(* Logix 5000 project; controller CIP_14485201 vendor 1 type 14 code 216 rev 38.11; software revision 38.01; part 4 of 12 *)
(* tags used below, declared in another part *)
   Alarm_Ack : INT[8];   // ALARMS ACKNOWLEDGE BITS
   Alarm_Present : INT[8];   // ALARM MSGS 1-127 PRESENT BITS
   Alarm_Remote_Ack_All : BOOL;   // SYSTEM ALARM ACK ALL TAG USED ON ALARM SETUP ADVANCED TAB TOGGLES EVEYTIME THE ACK_ALL BUTTON IS PUSHED
   Alarm_Timer : TIMER[128];   // ALARM MSGS 1-127 DELAY TIMERS
   Bit : BOOL[128];   // BIT
   IO_Status : INT;   // REMOTE I/O STATUS
   IO_Status_Masked : INT;   // REMOTE I/O STATUS MASK
   OpCode_Pin : DINT[5];   // OPCODE PIN ARRAY
   Process_Heartbeat_Memory : BOOL;
   Process_to_CIP : Process_to_CIP;   // PROCESS SIGNALS TO CIP
   Recipe : RECIPE[41];   // RECIPES
   SCLD_DrainValve_Feedback : SCALE;   // DRAIN FLOW FEEDBACK POSITION 0-100%
   SCLD_Supply_Flow : SCALE;   // SUPPLY FLOW 0-60 GPM
   SCLD_Supply_Press : SCALE;   // SUPPLY PRESSURE 0-100 PSIG
   SCLD_Supply_Temp : SCALE;   // SUPPLY TEMPERATURE 0-100°C
   SCLD_SupplyValve_Feedback : SCALE;   // SUPPLY FLOW FEEDBACK POSITION 0-100%
   SP_DrainValve_HighDeadband : REAL;   // CURRENT DRAIN VALVE DEADBAND SETPOINT
   SP_DrainValve_LowDeadband : REAL;   // CURRENT DRAIN VALVE DEADBAND SETPOINT
   SP_SupplyValve_HighDeadband : REAL;   // CURRENT SUPPLY VALVE DEADBAND SETPOINT
   SP_SupplyValve_LowDeadband : REAL;   // CURRENT SUPPLY VALVE DEADBAND SETPOINT
   Timer : TIMER[99];   // TIMER
   Timer_Chem1_Pump : TIMER[7];   // CHEM #1 CONTROL TIMERS
   Timer_Chem2_Pump : TIMER[7];   // CHEM #2 CONTROL TIMERS
(* MainProgram, continued *)

ROUTINE _05_ALARMS   (* ladder *)
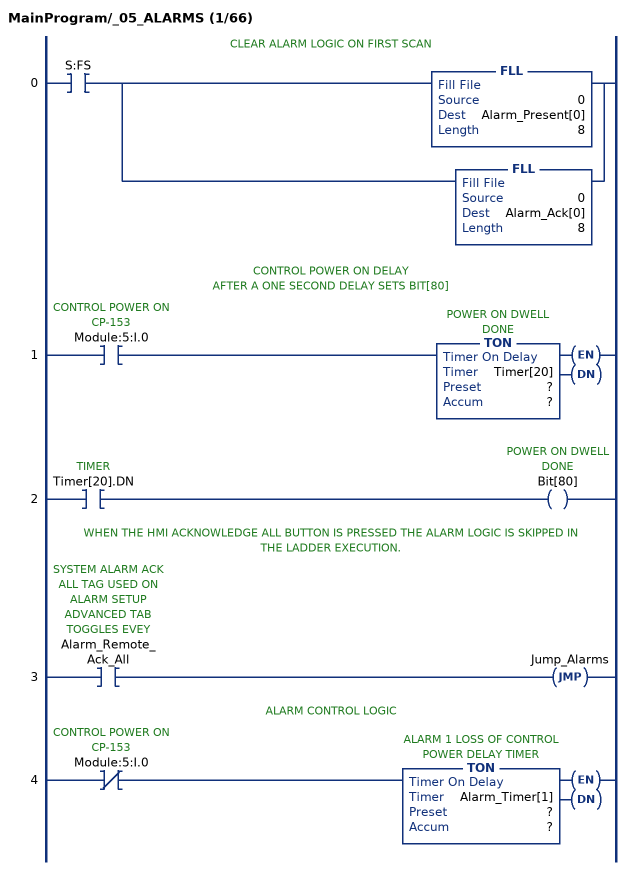
   // CLEAR ALARM LOGIC ON FIRST SCAN
   0: XIC(S:FS)[FLL(0,Alarm_Present[0],8) ,FLL(0,Alarm_Ack[0],8) ];
   // CONTROL POWER ON DELAY
   // AFTER A ONE SECOND DELAY SETS BIT[80]
   1: XIC(Module:5:I.0)TON(Timer[20],?,?);
   2: XIC(Timer[20].DN)OTE(Bit[80]);
   // WHEN THE HMI ACKNOWLEDGE ALL BUTTON IS PRESSED THE ALARM LOGIC IS SKIPPED IN THE LADDER EXECUTION.
   3: XIC(Alarm_Remote_Ack_All)JMP(Jump_Alarms);
   // ALARM CONTROL LOGIC
   4: XIO(Module:5:I.0)TON(Alarm_Timer[1],?,?);
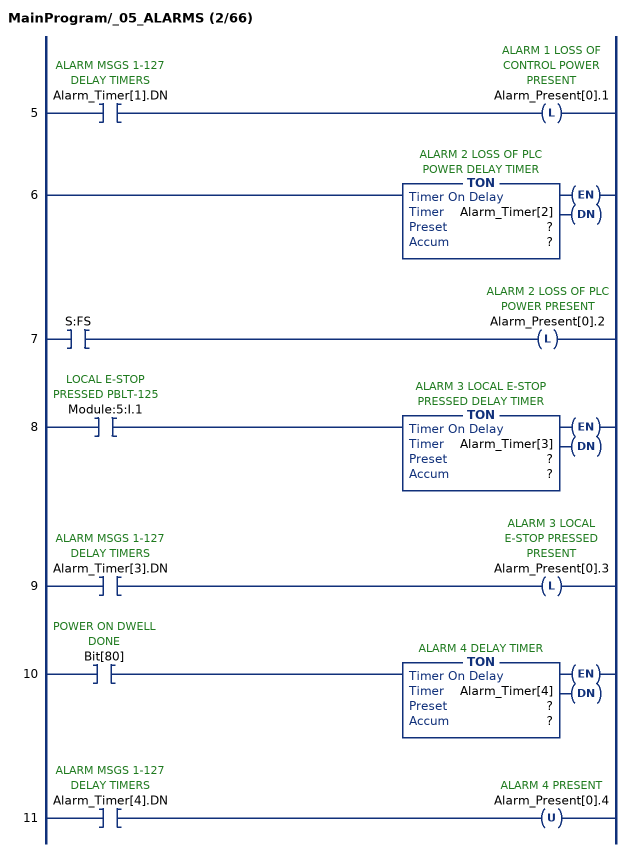
   5: XIC(Alarm_Timer[1].DN)OTL(Alarm_Present[0].1);
   6: TON(Alarm_Timer[2],?,?);
   7: XIC(S:FS)OTL(Alarm_Present[0].2);
   8: XIC(Module:5:I.1)TON(Alarm_Timer[3],?,?);
   9: XIC(Alarm_Timer[3].DN)OTL(Alarm_Present[0].3);
   10: XIC(Bit[80])TON(Alarm_Timer[4],?,?);
   11: XIC(Alarm_Timer[4].DN)OTU(Alarm_Present[0].4);
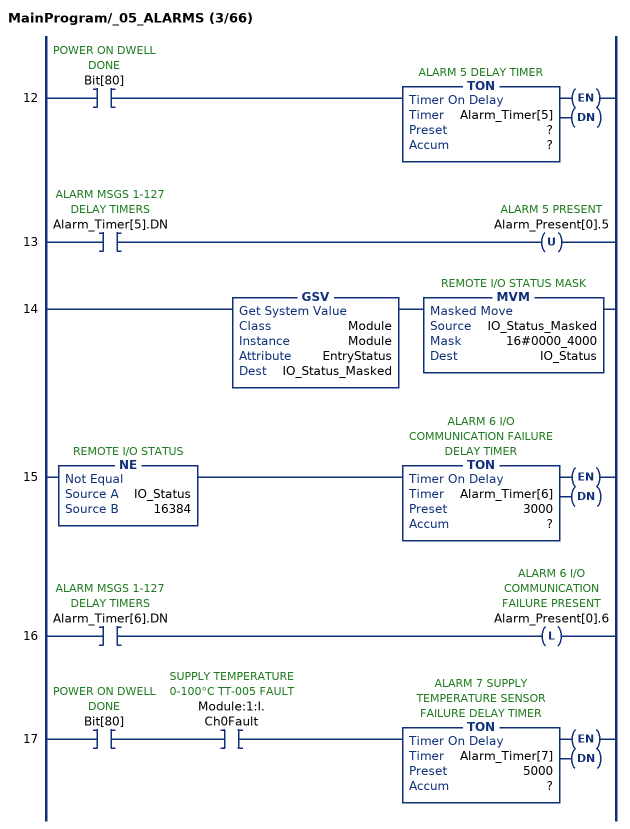
   12: XIC(Bit[80])TON(Alarm_Timer[5],?,?);
   13: XIC(Alarm_Timer[5].DN)OTU(Alarm_Present[0].5);
   14: GSV(Module,Module,EntryStatus,IO_Status_Masked)MVM(IO_Status_Masked,16#0000_4000,IO_Status);
   15: NE(IO_Status,16384)TON(Alarm_Timer[6],?,?);
   16: XIC(Alarm_Timer[6].DN)OTL(Alarm_Present[0].6);
   17: XIC(Bit[80])XIC(Module:1:I.Ch0Fault)TON(Alarm_Timer[7],?,?);
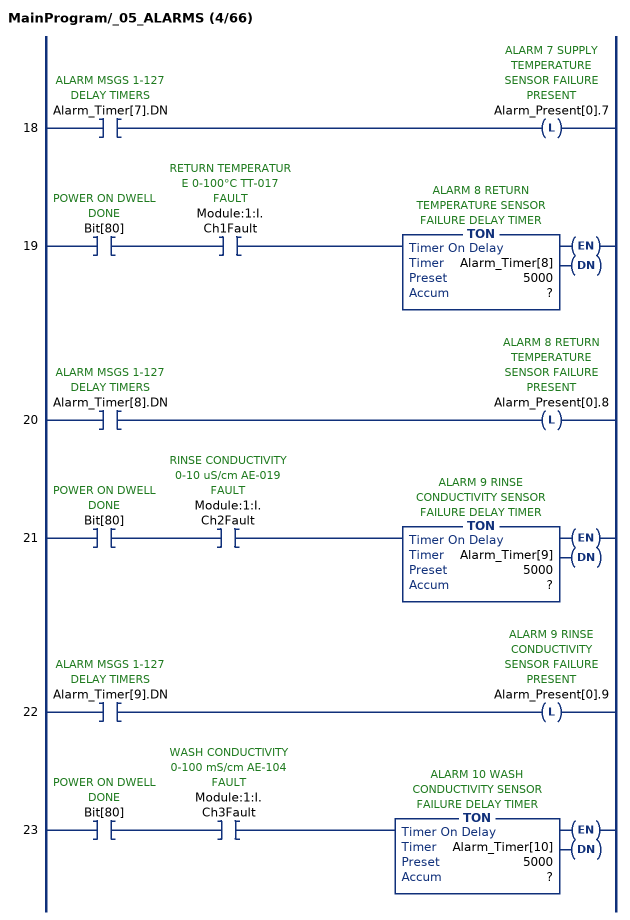
   18: XIC(Alarm_Timer[7].DN)OTL(Alarm_Present[0].7);
   19: XIC(Bit[80])XIC(Module:1:I.Ch1Fault)TON(Alarm_Timer[8],?,?);
   20: XIC(Alarm_Timer[8].DN)OTL(Alarm_Present[0].8);
   21: XIC(Bit[80])XIC(Module:1:I.Ch2Fault)TON(Alarm_Timer[9],?,?);
   22: XIC(Alarm_Timer[9].DN)OTL(Alarm_Present[0].9);
   23: XIC(Bit[80])XIC(Module:1:I.Ch3Fault)TON(Alarm_Timer[10],?,?);
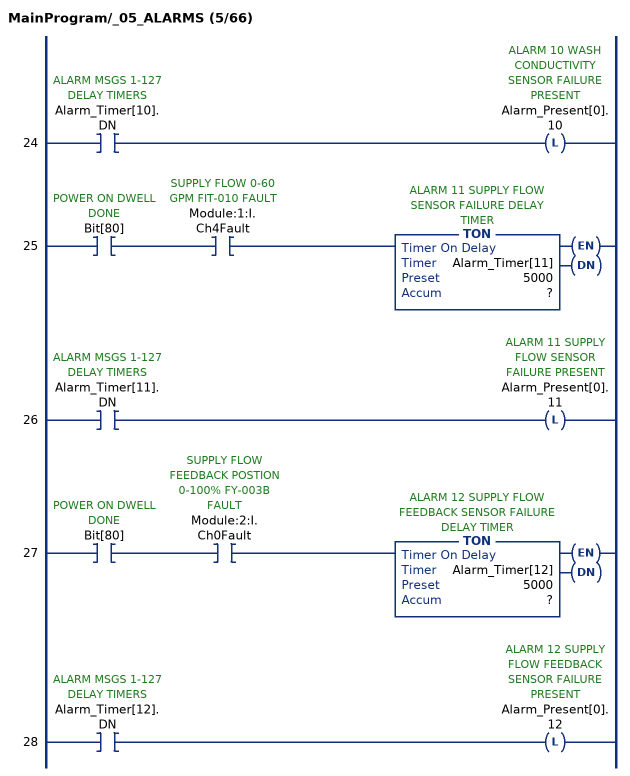
   24: XIC(Alarm_Timer[10].DN)OTL(Alarm_Present[0].10);
   25: XIC(Bit[80])XIC(Module:1:I.Ch4Fault)TON(Alarm_Timer[11],?,?);
   26: XIC(Alarm_Timer[11].DN)OTL(Alarm_Present[0].11);
   27: XIC(Bit[80])XIC(Module:2:I.Ch0Fault)TON(Alarm_Timer[12],?,?);
   28: XIC(Alarm_Timer[12].DN)OTL(Alarm_Present[0].12);
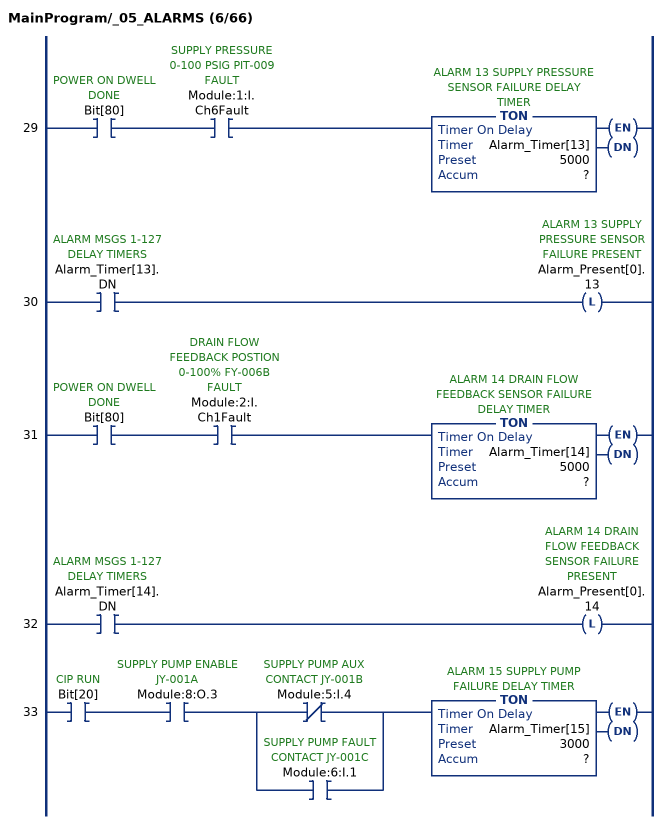
   29: XIC(Bit[80])XIC(Module:1:I.Ch6Fault)TON(Alarm_Timer[13],?,?);
   30: XIC(Alarm_Timer[13].DN)OTL(Alarm_Present[0].13);
   31: XIC(Bit[80])XIC(Module:2:I.Ch1Fault)TON(Alarm_Timer[14],?,?);
   32: XIC(Alarm_Timer[14].DN)OTL(Alarm_Present[0].14);
   33: XIC(Bit[20])XIC(Module:8:O.3)[XIO(Module:5:I.4) ,XIC(Module:6:I.1) ]TON(Alarm_Timer[15],?,?);
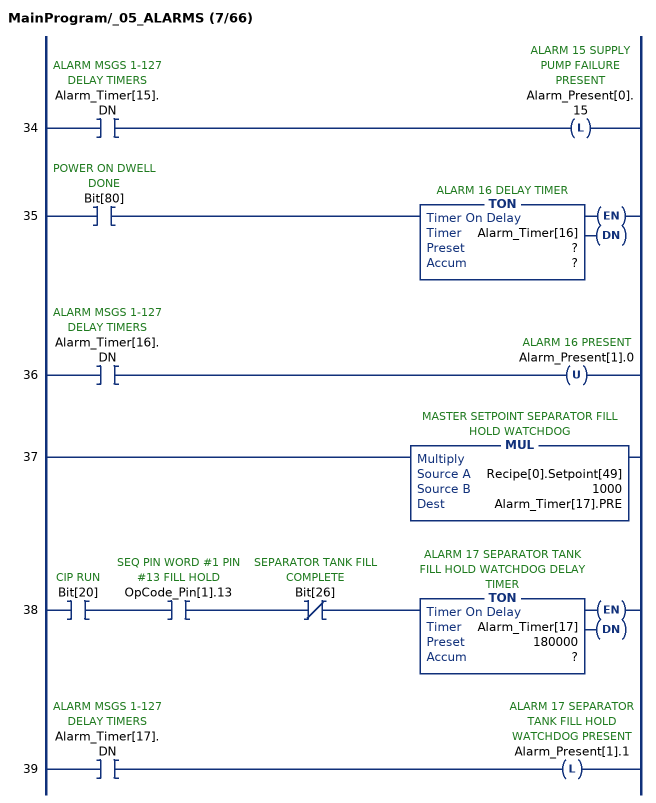
   34: XIC(Alarm_Timer[15].DN)OTL(Alarm_Present[0].15);
   35: XIC(Bit[80])TON(Alarm_Timer[16],?,?);
   36: XIC(Alarm_Timer[16].DN)OTU(Alarm_Present[1].0);
   37: MUL(Recipe[0].Setpoint[49],1000,Alarm_Timer[17].PRE);
   38: XIC(Bit[20])XIC(OpCode_Pin[1].13)XIO(Bit[26])TON(Alarm_Timer[17],?,?);
   39: XIC(Alarm_Timer[17].DN)OTL(Alarm_Present[1].1);
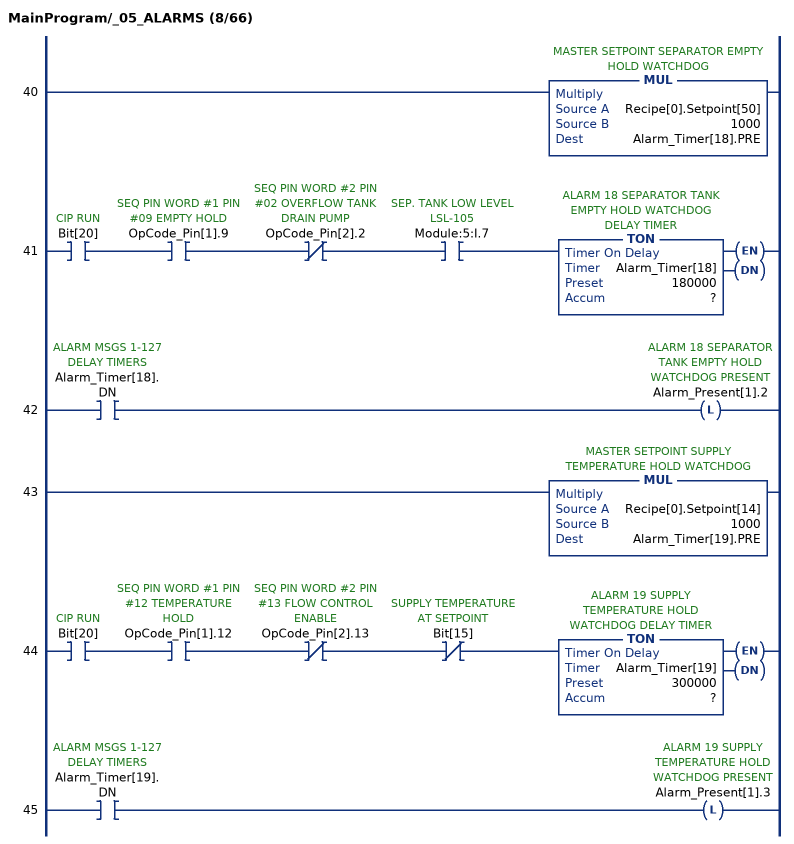
   40: MUL(Recipe[0].Setpoint[50],1000,Alarm_Timer[18].PRE);
   41: XIC(Bit[20])XIC(OpCode_Pin[1].9)XIO(OpCode_Pin[2].2)XIC(Module:5:I.7)TON(Alarm_Timer[18],?,?);
   42: XIC(Alarm_Timer[18].DN)OTL(Alarm_Present[1].2);
   43: MUL(Recipe[0].Setpoint[14],1000,Alarm_Timer[19].PRE);
   44: XIC(Bit[20])XIC(OpCode_Pin[1].12)XIO(OpCode_Pin[2].13)XIO(Bit[15])TON(Alarm_Timer[19],?,?);
   45: XIC(Alarm_Timer[19].DN)OTL(Alarm_Present[1].3);
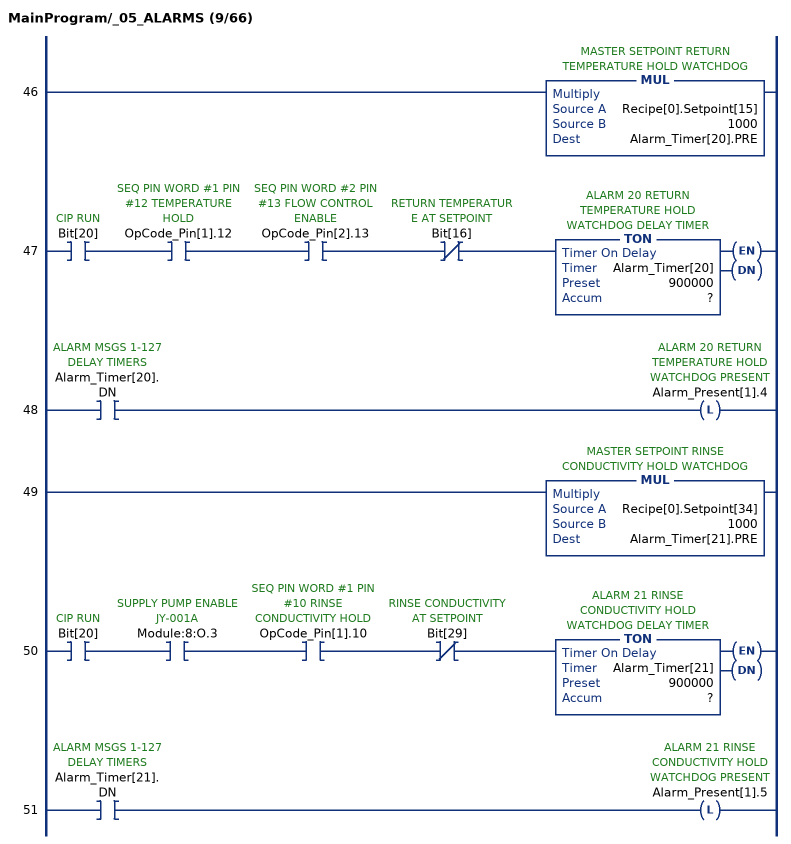
   46: MUL(Recipe[0].Setpoint[15],1000,Alarm_Timer[20].PRE);
   47: XIC(Bit[20])XIC(OpCode_Pin[1].12)XIC(OpCode_Pin[2].13)XIO(Bit[16])TON(Alarm_Timer[20],?,?);
   48: XIC(Alarm_Timer[20].DN)OTL(Alarm_Present[1].4);
   49: MUL(Recipe[0].Setpoint[34],1000,Alarm_Timer[21].PRE);
   50: XIC(Bit[20])XIC(Module:8:O.3)XIC(OpCode_Pin[1].10)XIO(Bit[29])TON(Alarm_Timer[21],?,?);
   51: XIC(Alarm_Timer[21].DN)OTL(Alarm_Present[1].5);
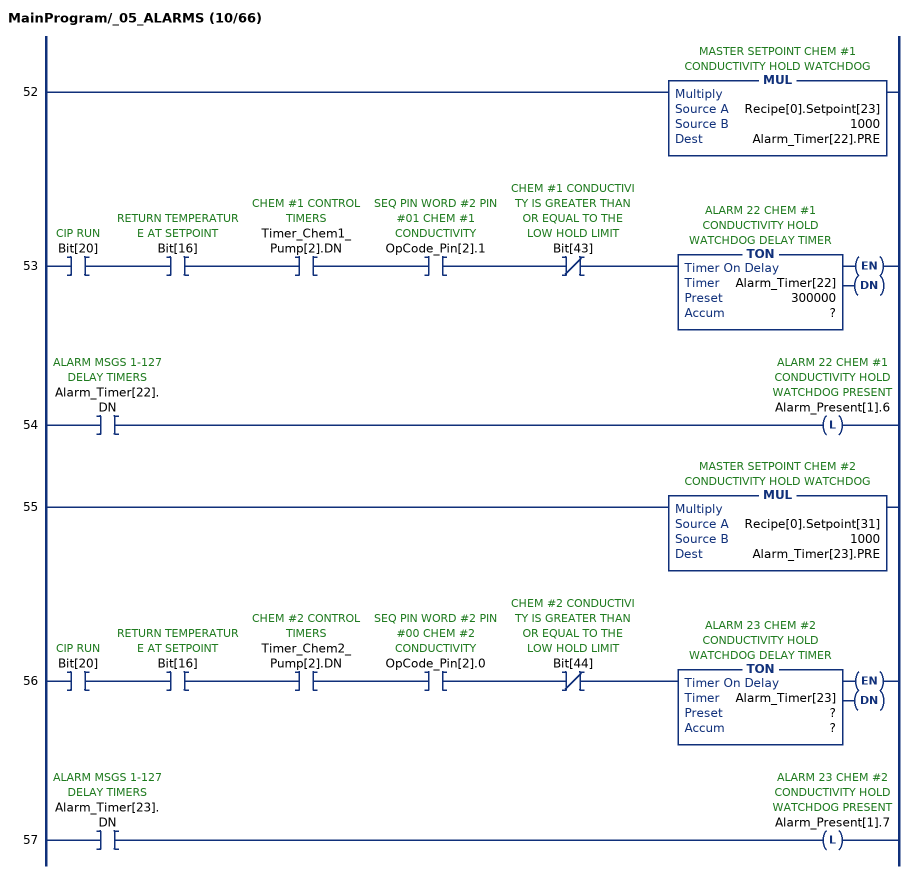
   52: MUL(Recipe[0].Setpoint[23],1000,Alarm_Timer[22].PRE);
   53: XIC(Bit[20])XIC(Bit[16])XIC(Timer_Chem1_Pump[2].DN)XIC(OpCode_Pin[2].1)XIO(Bit[43])TON(Alarm_Timer[22],?,?);
   54: XIC(Alarm_Timer[22].DN)OTL(Alarm_Present[1].6);
   55: MUL(Recipe[0].Setpoint[31],1000,Alarm_Timer[23].PRE);
   56: XIC(Bit[20])XIC(Bit[16])XIC(Timer_Chem2_Pump[2].DN)XIC(OpCode_Pin[2].0)XIO(Bit[44])TON(Alarm_Timer[23],?,?);
   57: XIC(Alarm_Timer[23].DN)OTL(Alarm_Present[1].7);
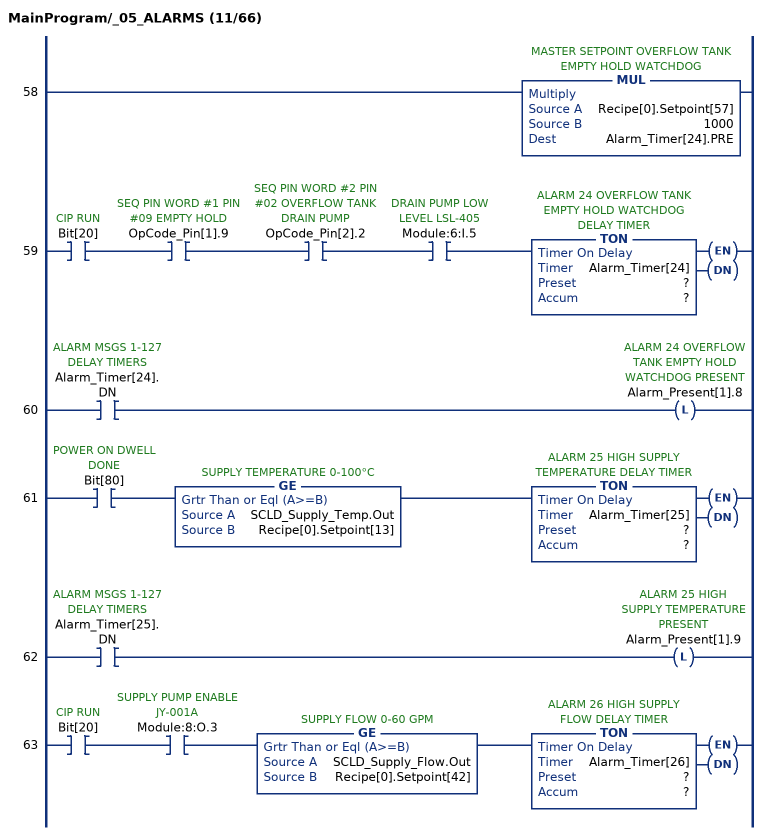
   58: MUL(Recipe[0].Setpoint[57],1000,Alarm_Timer[24].PRE);
   59: XIC(Bit[20])XIC(OpCode_Pin[1].9)XIC(OpCode_Pin[2].2)XIC(Module:6:I.5)TON(Alarm_Timer[24],?,?);
   60: XIC(Alarm_Timer[24].DN)OTL(Alarm_Present[1].8);
   61: XIC(Bit[80])GE(SCLD_Supply_Temp.Out,Recipe[0].Setpoint[13])TON(Alarm_Timer[25],?,?);
   62: XIC(Alarm_Timer[25].DN)OTL(Alarm_Present[1].9);
   63: XIC(Bit[20])XIC(Module:8:O.3)GE(SCLD_Supply_Flow.Out,Recipe[0].Setpoint[42])TON(Alarm_Timer[26],?,?);
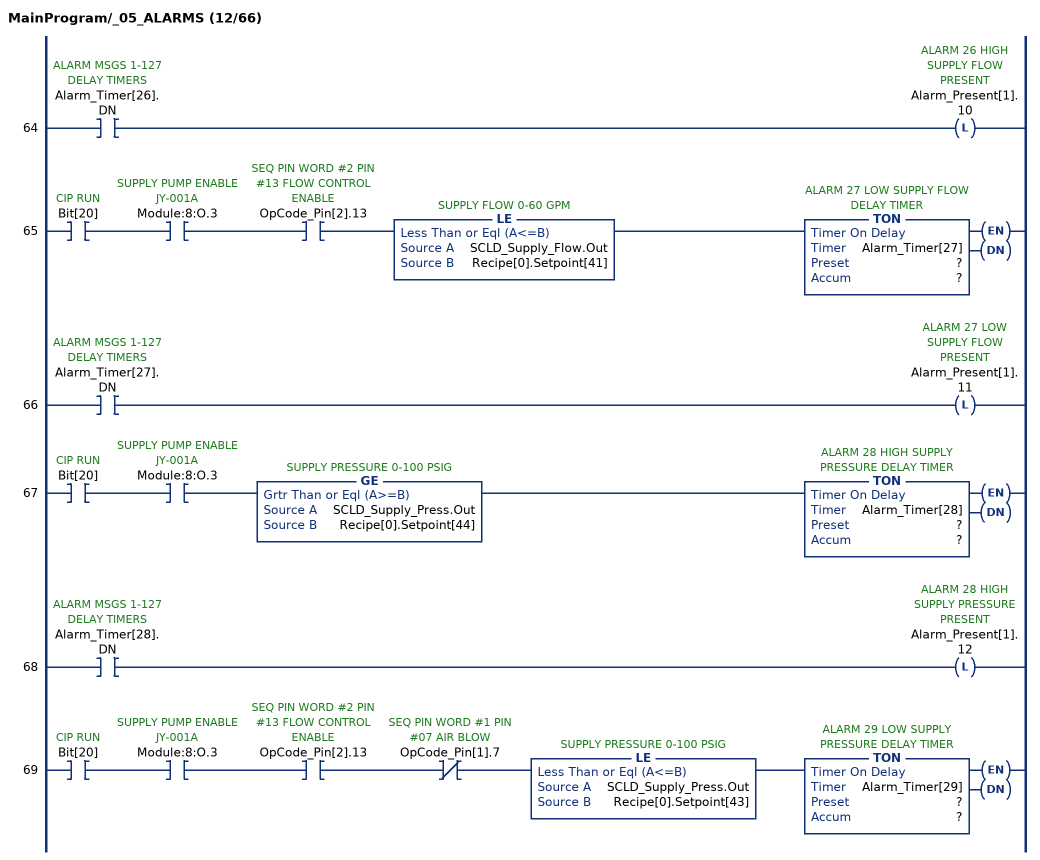
   64: XIC(Alarm_Timer[26].DN)OTL(Alarm_Present[1].10);
   65: XIC(Bit[20])XIC(Module:8:O.3)XIC(OpCode_Pin[2].13)LE(SCLD_Supply_Flow.Out,Recipe[0].Setpoint[41])TON(Alarm_Timer[27],?,?);
   66: XIC(Alarm_Timer[27].DN)OTL(Alarm_Present[1].11);
   67: XIC(Bit[20])XIC(Module:8:O.3)GE(SCLD_Supply_Press.Out,Recipe[0].Setpoint[44])TON(Alarm_Timer[28],?,?);
   68: XIC(Alarm_Timer[28].DN)OTL(Alarm_Present[1].12);
   69: XIC(Bit[20])XIC(Module:8:O.3)XIC(OpCode_Pin[2].13)XIO(OpCode_Pin[1].7)LE(SCLD_Supply_Press.Out,Recipe[0].Setpoint[43])TON(Alarm_Timer[29],?,?);
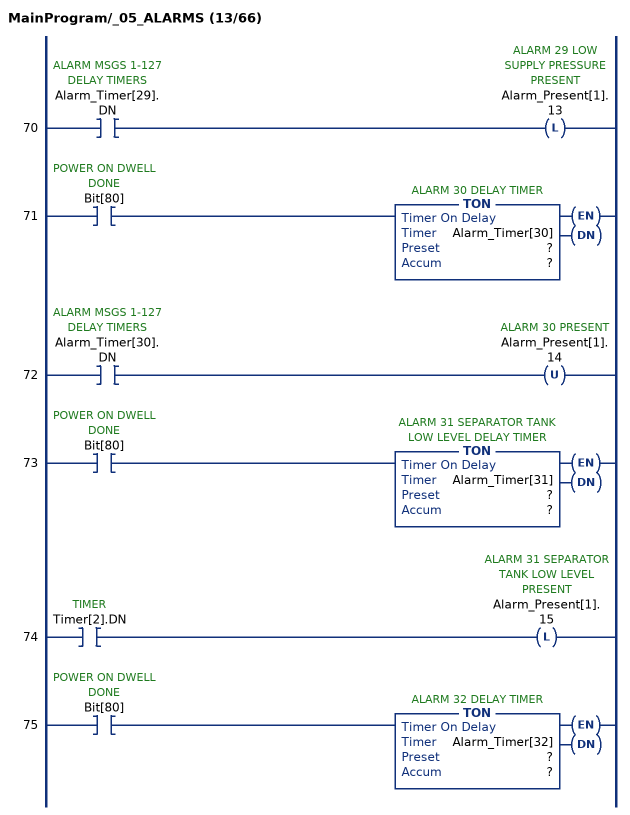
   70: XIC(Alarm_Timer[29].DN)OTL(Alarm_Present[1].13);
   71: XIC(Bit[80])TON(Alarm_Timer[30],?,?);
   72: XIC(Alarm_Timer[30].DN)OTU(Alarm_Present[1].14);
   73: XIC(Bit[80])TON(Alarm_Timer[31],?,?);
   74: XIC(Timer[2].DN)OTL(Alarm_Present[1].15);
   75: XIC(Bit[80])TON(Alarm_Timer[32],?,?);
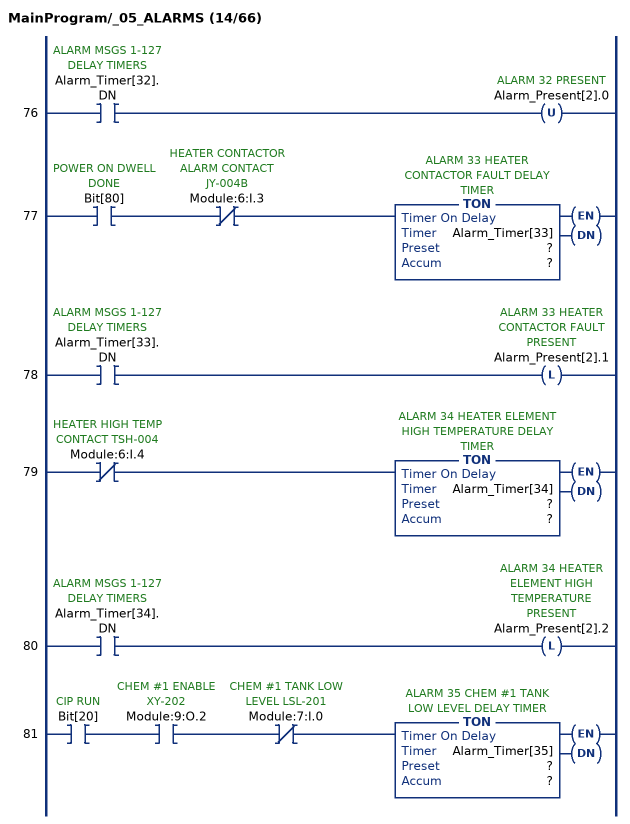
   76: XIC(Alarm_Timer[32].DN)OTU(Alarm_Present[2].0);
   77: XIC(Bit[80])XIO(Module:6:I.3)TON(Alarm_Timer[33],?,?);
   78: XIC(Alarm_Timer[33].DN)OTL(Alarm_Present[2].1);
   79: XIO(Module:6:I.4)TON(Alarm_Timer[34],?,?);
   80: XIC(Alarm_Timer[34].DN)OTL(Alarm_Present[2].2);
   81: XIC(Bit[20])XIC(Module:9:O.2)XIO(Module:7:I.0)TON(Alarm_Timer[35],?,?);
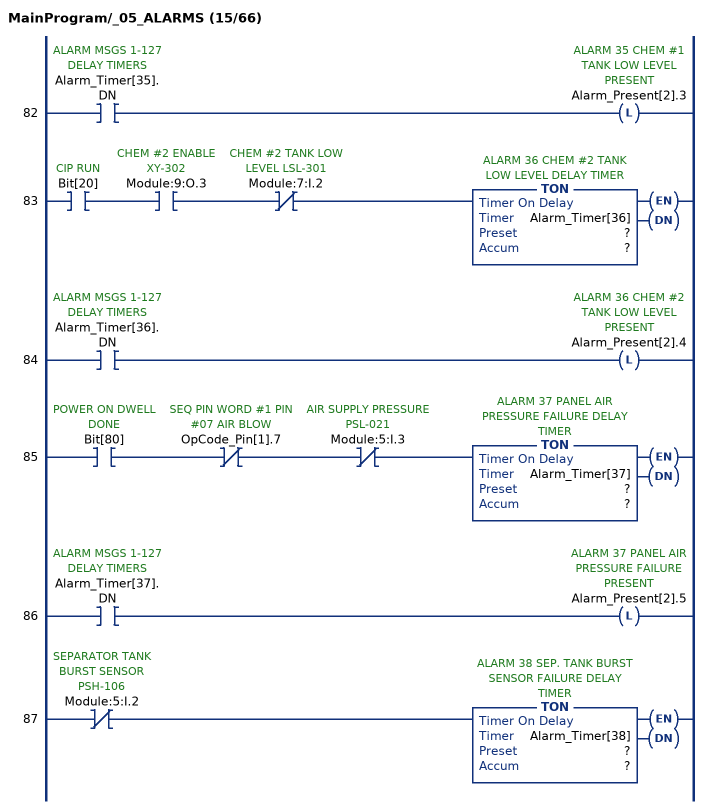
   82: XIC(Alarm_Timer[35].DN)OTL(Alarm_Present[2].3);
   83: XIC(Bit[20])XIC(Module:9:O.3)XIO(Module:7:I.2)TON(Alarm_Timer[36],?,?);
   84: XIC(Alarm_Timer[36].DN)OTL(Alarm_Present[2].4);
   85: XIC(Bit[80])XIO(OpCode_Pin[1].7)XIO(Module:5:I.3)TON(Alarm_Timer[37],?,?);
   86: XIC(Alarm_Timer[37].DN)OTL(Alarm_Present[2].5);
   87: XIO(Module:5:I.2)TON(Alarm_Timer[38],?,?);
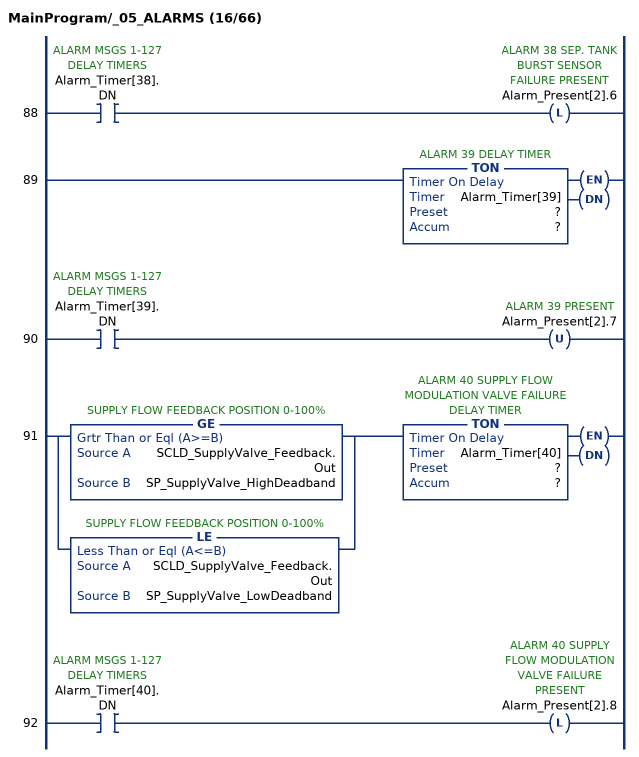
   88: XIC(Alarm_Timer[38].DN)OTL(Alarm_Present[2].6);
   89: TON(Alarm_Timer[39],?,?);
   90: XIC(Alarm_Timer[39].DN)OTU(Alarm_Present[2].7);
   91: [GE(SCLD_SupplyValve_Feedback.Out,SP_SupplyValve_HighDeadband) ,LE(SCLD_SupplyValve_Feedback.Out,SP_SupplyValve_LowDeadband) ]TON(Alarm_Timer[40],?,?);
   92: XIC(Alarm_Timer[40].DN)OTL(Alarm_Present[2].8);
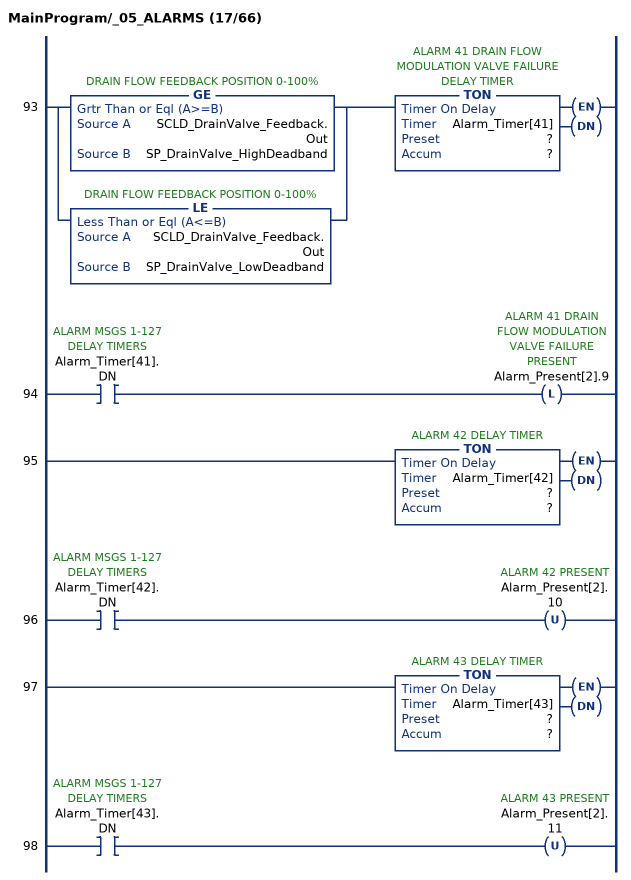
   93: [GE(SCLD_DrainValve_Feedback.Out,SP_DrainValve_HighDeadband) ,LE(SCLD_DrainValve_Feedback.Out,SP_DrainValve_LowDeadband) ]TON(Alarm_Timer[41],?,?);
   94: XIC(Alarm_Timer[41].DN)OTL(Alarm_Present[2].9);
   95: TON(Alarm_Timer[42],?,?);
   96: XIC(Alarm_Timer[42].DN)OTU(Alarm_Present[2].10);
   97: TON(Alarm_Timer[43],?,?);
   98: XIC(Alarm_Timer[43].DN)OTU(Alarm_Present[2].11);
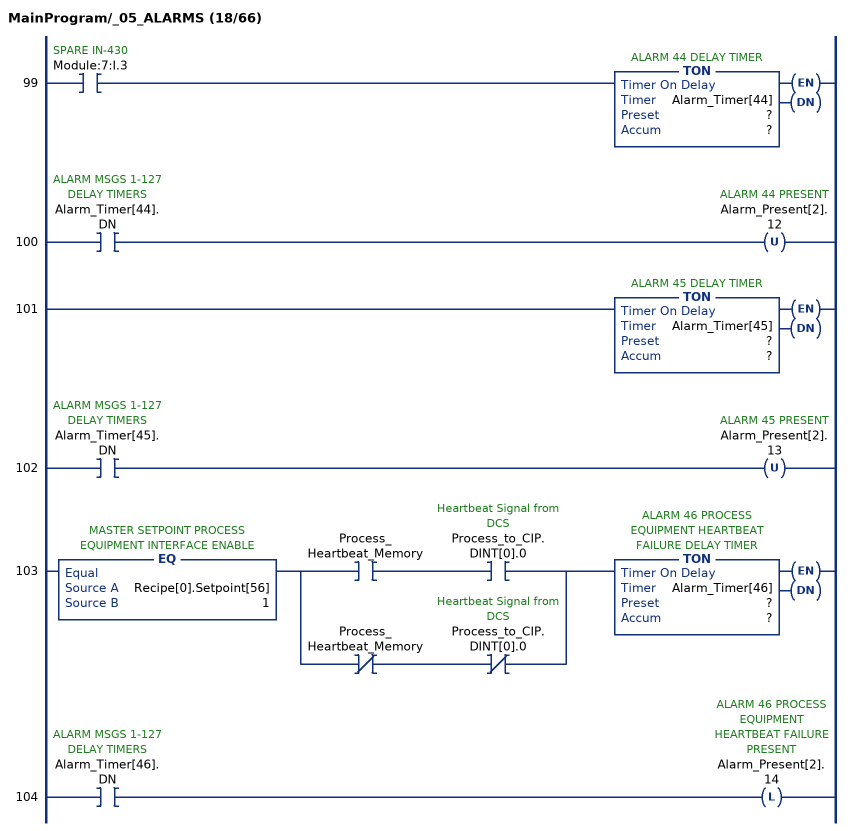
   99: XIC(Module:7:I.3)TON(Alarm_Timer[44],?,?);
   100: XIC(Alarm_Timer[44].DN)OTU(Alarm_Present[2].12);
   101: TON(Alarm_Timer[45],?,?);
   102: XIC(Alarm_Timer[45].DN)OTU(Alarm_Present[2].13);
   103: EQ(Recipe[0].Setpoint[56],1)[XIC(Process_Heartbeat_Memory) XIC(Process_to_CIP.DINT[0].0) ,XIO(Process_Heartbeat_Memory) XIO(Process_to_CIP.DINT[0].0) ]TON(Alarm_Timer[46],?,?);
   104: XIC(Alarm_Timer[46].DN)OTL(Alarm_Present[2].14);
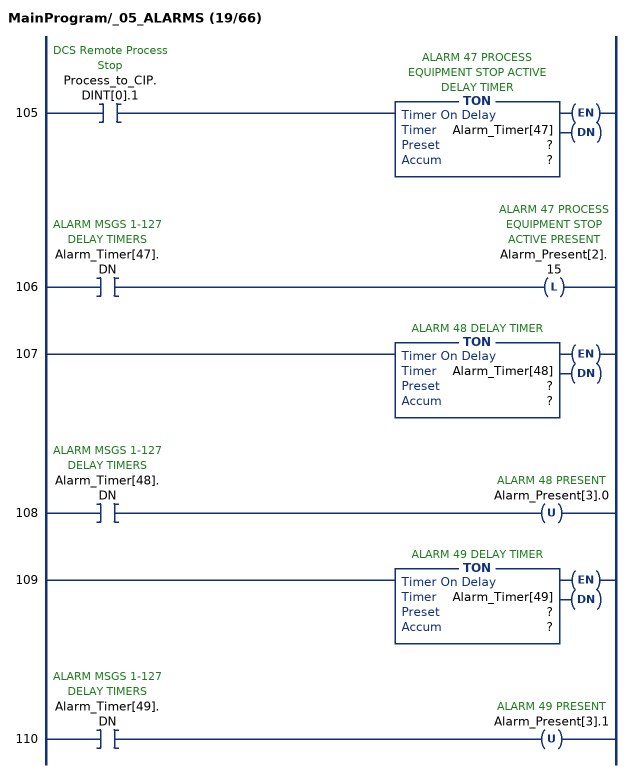
   105: XIC(Process_to_CIP.DINT[0].1)TON(Alarm_Timer[47],?,?);
   106: XIC(Alarm_Timer[47].DN)OTL(Alarm_Present[2].15);
   107: TON(Alarm_Timer[48],?,?);
   108: XIC(Alarm_Timer[48].DN)OTU(Alarm_Present[3].0);
   109: TON(Alarm_Timer[49],?,?);
   110: XIC(Alarm_Timer[49].DN)OTU(Alarm_Present[3].1);
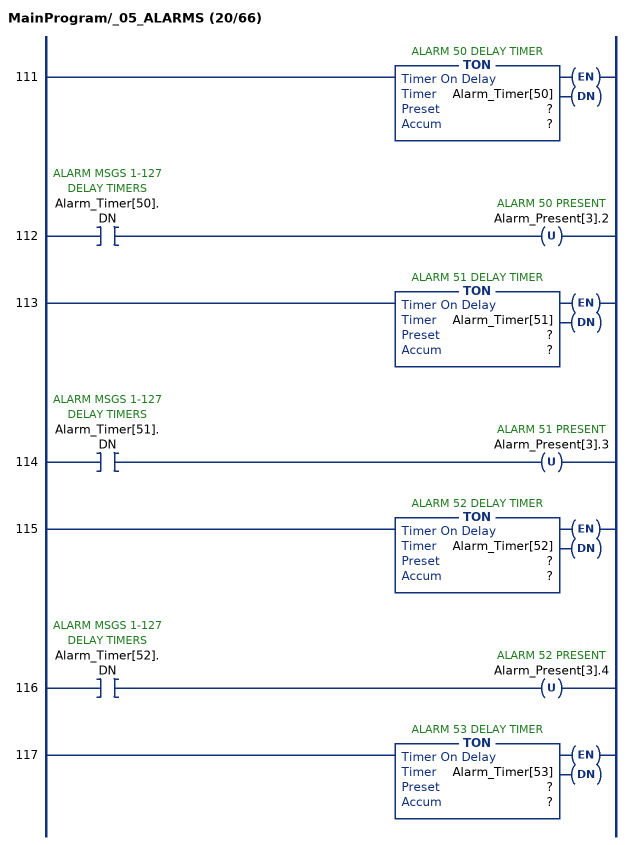
   111: TON(Alarm_Timer[50],?,?);
   112: XIC(Alarm_Timer[50].DN)OTU(Alarm_Present[3].2);
   113: TON(Alarm_Timer[51],?,?);
   114: XIC(Alarm_Timer[51].DN)OTU(Alarm_Present[3].3);
   115: TON(Alarm_Timer[52],?,?);
   116: XIC(Alarm_Timer[52].DN)OTU(Alarm_Present[3].4);
   117: TON(Alarm_Timer[53],?,?);
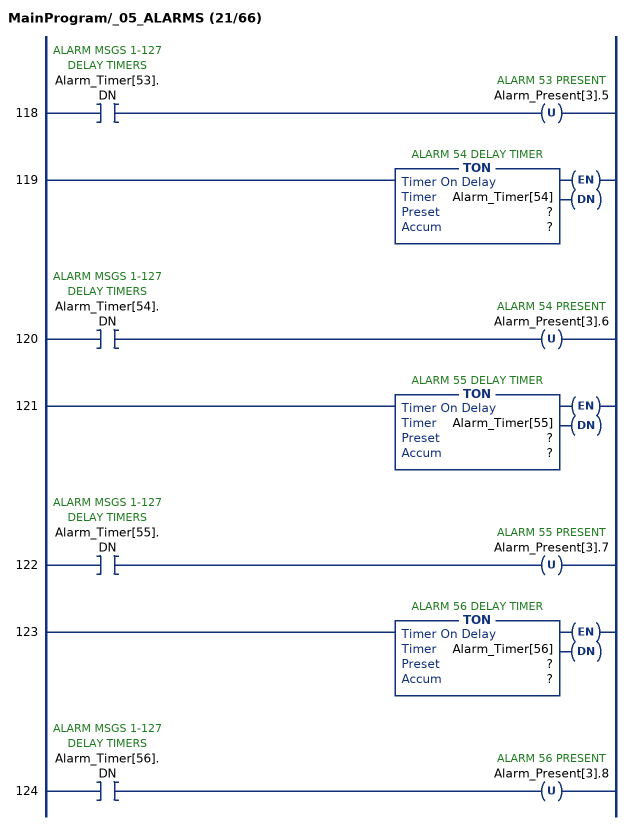
   118: XIC(Alarm_Timer[53].DN)OTU(Alarm_Present[3].5);
   119: TON(Alarm_Timer[54],?,?);
   120: XIC(Alarm_Timer[54].DN)OTU(Alarm_Present[3].6);
   121: TON(Alarm_Timer[55],?,?);
   122: XIC(Alarm_Timer[55].DN)OTU(Alarm_Present[3].7);
   123: TON(Alarm_Timer[56],?,?);
   124: XIC(Alarm_Timer[56].DN)OTU(Alarm_Present[3].8);
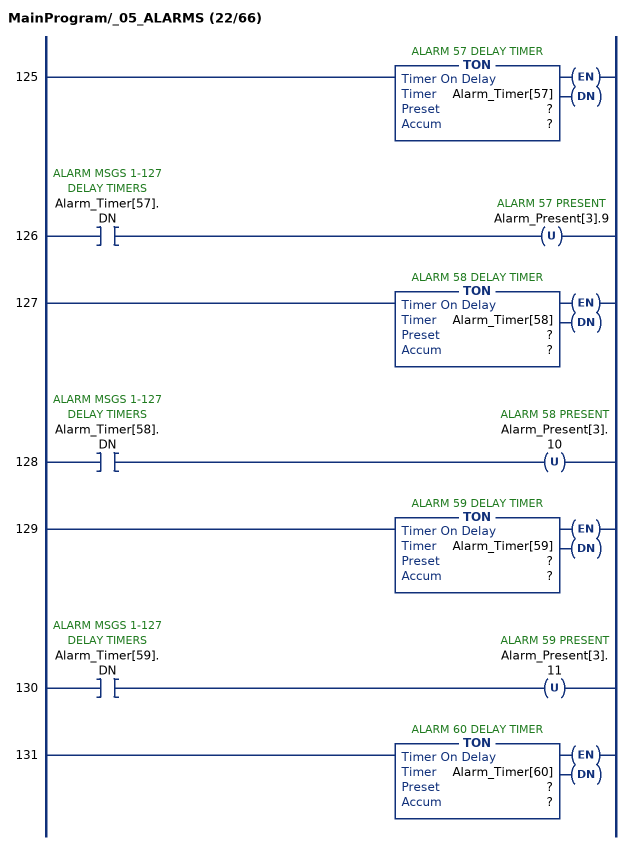
   125: TON(Alarm_Timer[57],?,?);
   126: XIC(Alarm_Timer[57].DN)OTU(Alarm_Present[3].9);
   127: TON(Alarm_Timer[58],?,?);
   128: XIC(Alarm_Timer[58].DN)OTU(Alarm_Present[3].10);
   129: TON(Alarm_Timer[59],?,?);
   130: XIC(Alarm_Timer[59].DN)OTU(Alarm_Present[3].11);
   131: TON(Alarm_Timer[60],?,?);
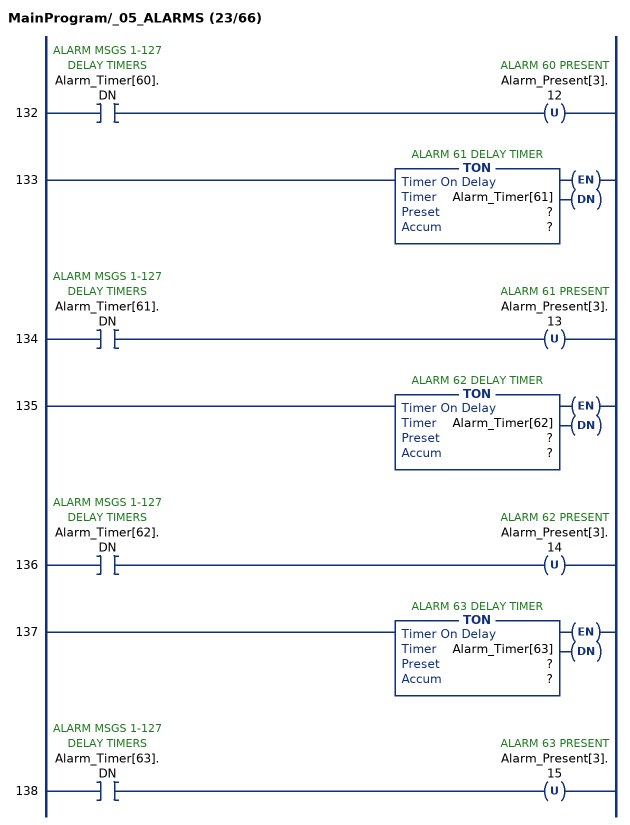
   132: XIC(Alarm_Timer[60].DN)OTU(Alarm_Present[3].12);
   133: TON(Alarm_Timer[61],?,?);
   134: XIC(Alarm_Timer[61].DN)OTU(Alarm_Present[3].13);
   135: TON(Alarm_Timer[62],?,?);
   136: XIC(Alarm_Timer[62].DN)OTU(Alarm_Present[3].14);
   137: TON(Alarm_Timer[63],?,?);
   138: XIC(Alarm_Timer[63].DN)OTU(Alarm_Present[3].15);
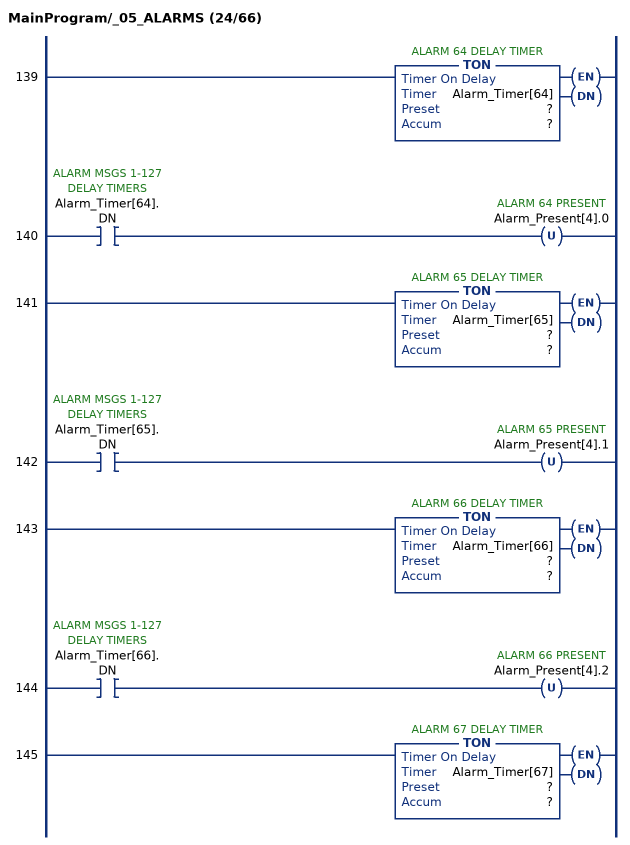
   139: TON(Alarm_Timer[64],?,?);
   140: XIC(Alarm_Timer[64].DN)OTU(Alarm_Present[4].0);
   141: TON(Alarm_Timer[65],?,?);
   142: XIC(Alarm_Timer[65].DN)OTU(Alarm_Present[4].1);
   143: TON(Alarm_Timer[66],?,?);
   144: XIC(Alarm_Timer[66].DN)OTU(Alarm_Present[4].2);
   145: TON(Alarm_Timer[67],?,?);
